Fanuc KAREL source: KT00976.KL

PROGRAM KT00976
%NOLOCKGROUP
VAR
  ENTRY: INTEGER
  PNAME: STRING[80]
  VNAME: STRING[80]
  STATUS: INTEGER
  VALUE: ARRAY[4] OF JOINTPOS
BEGIN
  ENTRY = 0
  PNAME = ''
  VNAME = 'VALUE'
  SET_VAR(ENTRY, PNAME, VNAME, VALUE, STATUS)
END KT00976
